DATA_BLOCK "GDB_SequenceHelperTest"
{ S7_Optimized_Access := 'TRUE' }
VERSION : 0.1
NON_RETAIN
VAR
    Seq {ExternalWritable := 'False'} : "FRK_SequenceCtx";
    Row {ExternalWritable := 'False'} : "FRK_SequenceRow";
    Diag : "ST_Diagnostic";
    WaitOk {ExternalWritable := 'False'} : Bool;
END_VAR
BEGIN
END_DATA_BLOCK
